FUNCTION F_iFB_Num_sFB_Num : STRING(3)
VAR_INPUT
	iFB_Num: INT;
END_VAR
VAR
END_VAR

IF iFB_Num<10 THEN;
	F_iFB_Num_sFB_Num:=CONCAT(STR1:='00',STR2:=INT_TO_STRING(iFB_Num));
ELSIF iFB_Num<100 THEN;
	F_iFB_Num_sFB_Num:=CONCAT(STR1:='0',STR2:=INT_TO_STRING(iFB_Num));
ELSE;
	F_iFB_Num_sFB_Num:=CONCAT(STR1:='',STR2:=INT_TO_STRING(iFB_Num));
END_IF

END_FUNCTION

(* stored: Version 1.1.0.1, ProductVersion 3.1.4024.13
   POU F_iFB_Num_sFB_Num: Id {0fc1480b-3d38-49c4-85cc-de6fbc710349}, SpecialFunc None *)
